FUNCTION F_JsonInt : BOOL
VAR_INPUT
    sKey   : STRING(31);
    nValue : DINT;
END_VAR
VAR_IN_OUT
    fbJson : FB_JsonSaxWriter;
END_VAR

fbJson.AddKey(sKey);
fbJson.AddDint(nValue);
F_JsonInt := TRUE;

END_FUNCTION

(* stored: Version 1.1.0.1
   POU F_JsonInt: Id {696ba799-6306-4e45-9a59-ed9d08410e72}, SpecialFunc None *)
